(* IEC 61131-3 sources: JingjiangArm/moonboxpro_arm_8.4/Application/Application/任务列表/ExtTask/动作处理/工艺辅助/冷风, 2 files *)

(* ---- KS_ReCfgCoolBlowerIO.st ---- *)
(*@CES
Name=KS_ReCfgCoolBlowerIO
Type=FunctionBlock
TypeGuid=6f9dac99-8de1-4efc-8465-68ac443b7d08
Guid=0f7b114d-d936-480a-be34-fd41a916f68a
HasDeclaration=True
HasImplementation=True
*)
{DECLARATION}
FUNCTION KS_ReCfgCoolBlowerIO : bool
VAR_INPUT
	i_xInput				: BOOL;(*输入重新分配*)
	i_xOutput				: BOOL;(*输出重新分配*)
	i_xCoolBlowerFlag		: BOOL;(*全体冷风启动标志*)
	i_iGrpAxisNum_Pu		:INT ;
	i_aiGrpAxisList			: ARRAY [1..MAX_UNIT_NUM] OF INT;(*系的轴列表*)
	i_paxAxisStartEn		: POINTER TO ARRAY [1..MAX_UNIT_NUM] OF BOOL;(*轴启动使能|有效后按钮开关才能起作用*)
	i_paxStartKnob			: POINTER TO ARRAY [1..MAX_UNIT_NUM] OF BOOL;(*全体启动,每个轴旋钮输入*)
	i_paxStartOrStopBtn		: POINTER TO ARRAY [1..MAX_UNIT_NUM] OF BOOL;(*单轴的启动停止按钮*)
	i_paxNeedStop			: POINTER TO ARRAY [1..MAX_UNIT_NUM] OF BOOL;(*单轴需要停止标志*)
	i_paxAxisStarted		: POINTER TO ARRAY [1..MAX_UNIT_NUM] OF BOOL;(*单个轴的启动输出标志|实际处于启动状态，																		可以根据i_paxNeedStop这个变量控制实际输出*)
	i_axCoolBlower			:ARRAY [1..MAX_UNIT_NUM] OF BOOL;
	i_axCoolBlower_Button			:ARRAY [1..MAX_UNIT_NUM] OF BOOL;
	i_paxLamp_CoolBlower			:POINTER TO ARRAY [1..MAX_UNIT_NUM] OF BOOL;
	i_paxRel_CoolBlower			:POINTER TO ARRAY [1..MAX_UNIT_NUM] OF BOOL;
	i_paxLamp_AllCoolBlower		:POINTER TO ARRAY [1..MAX_UNIT_NUM] OF BOOL;
	i_pxLamp_AllCoolBlower		: POINTER TO BOOL;

END_VAR
VAR_OUTPUT

END_VAR
VAR
	iUnitId: INT;
	iN: INT;
END_VAR

{IMPLEMENTATION}
IF i_paxAxisStartEn<>0 AND
	i_paxStartKnob<>0 AND
	i_paxNeedStop<>0 AND
 	i_paxStartOrStopBtn<>0 AND
	i_paxAxisStarted<>0  THEN
	IF i_xInput THEN
		FOR iN:=1 TO MAX_UNIT_NUM  BY 1 DO
			i_paxStartKnob^[iN]:=FALSE;
			i_paxStartOrStopBtn^[iN]:=FALSE;
			i_paxNeedStop^[iN]:=FALSE;
			i_paxAxisStartEn^[iN]:=FALSE;
		END_FOR

		FOR iN:=1 TO i_iGrpAxisNum_Pu  BY 1 DO
			iUnitId:=i_aiGrpAxisList[iN];
			IF iUnitId>0 AND iUnitId<= MAX_UNIT_NUM THEN
			i_paxStartKnob^[iUnitId]:=i_axCoolBlower[iUnitId];
			i_paxStartOrStopBtn^[iUnitId]:=i_axCoolBlower_Button[iUnitId];
			i_paxNeedStop^[iUnitId]:=FALSE;
			i_paxAxisStartEn^[iUnitId]:=TRUE; (*2024.3.14.165139*)
			END_IF
		END_FOR
	ELSIF i_xOutput THEN
		FOR iN:=1 TO i_iGrpAxisNum_Pu  BY 1 DO
			(*输出到牵引，*)

				iUnitId:=i_aiGrpAxisList[iN];
				IF iUnitId>0 AND iUnitId <= MAX_UNIT_NUM THEN(*输出循环到收牵，这样热风输出灯就可以配到收牵上了|2020.1.9.094955*)
					i_paxLamp_CoolBlower^[iUnitId]:=i_paxAxisStarted^[iUnitId];
					i_paxRel_CoolBlower^[iUnitId]:=i_paxAxisStarted^[iUnitId];
					i_paxLamp_AllCoolBlower^[iUnitId]:=i_xCoolBlowerFlag;
				END_IF

		END_FOR

	END_IF
END_IF

(* ---- KS_FB_GrpCoolBlowerCtrl.st ---- *)
(*@CES
Name=KS_FB_GrpCoolBlowerCtrl
Type=FunctionBlock
TypeGuid=6f9dac99-8de1-4efc-8465-68ac443b7d08
Guid=1cc9b71b-01ee-4c63-826f-1c195b3708a6
HasDeclaration=True
HasImplementation=True
*)
{DECLARATION}
FUNCTION_BLOCK KS_FB_GrpCoolBlowerCtrl
(*2020.10.14.090348重新处理*)
VAR_INPUT
	i_xEn: BOOL;
	i_iGrpId : INT;
	i_iAxisId_If: INT;
	i_iAxisId_Of: INT;
	i_iGrpAxisNum_Pu: INT; (*色组轴数*)
	i_aiGrpAxisList: ARRAY [1..MAX_UNIT_NUM] OF INT; (*系的轴列表*)
	i_pstStEvtReq:POINTER TO StEvtReq;
	i_xCoolBlowerByKnob:BOOL;(*单轴启动根据旋钮开关标志|用于全体开关控制启动的逻辑|无则不输入*)
	i_xStopCoolBlowerWhenEstop:BOOL;(*急停停止热风标志|有效了和急停关联，无效则不影响*)
	i_iCycleTime_Plc:INT;(*2024.01.22.142933+*)
	i_PastStIOMap_Axis_Extra_FE:  POINTER TO ARRAY [1..MAX_UNIT_NUM] OF StIOMap_Axis_Extra_FE  ;

	i_pastStIOMap_Main_FE	: POINTER TO ARRAY [1..4] OF StIOMap_Main_FE;(*轴io数据区域|*)
END_VAR
VAR_OUTPUT
	o_xEno: BOOL;
	o_iErNo: INT;(*0成功\-1参数无效|*)
	o_xCoolBlowerFlag:BOOL;
END_VAR
VAR
	fbKS_FB_CoolBlowerSys: KS_FB_BlowerFunction;
	axAxisStartKnob: ARRAY [1..MAX_UNIT_NUM] OF BOOL;
	axStartOrStopBtn: ARRAY [1..MAX_UNIT_NUM] OF BOOL;
	axNeedStop: ARRAY [1..MAX_UNIT_NUM] OF BOOL;
	axAxisStarted: ARRAY [1..MAX_UNIT_NUM] OF BOOL;
	axAxisStartEn: ARRAY [1..MAX_UNIT_NUM] OF BOOL;
	xCoolBlowerEn: BOOL;
	iStartedSum: INT;(*启动的轴数*)
	xFlag_Estop_In : BOOL;

	axCoolBlower_In			:ARRAY [1..MAX_UNIT_NUM] OF BOOL;
	axCoolBlower_Button_In			:ARRAY [1..MAX_UNIT_NUM] OF BOOL;

	xCoolBlower_In			: BOOL;
	xCoolBlower_Button_In			: BOOL;

	axLamp_CoolBlower_Out			: ARRAY [1..MAX_UNIT_NUM] OF BOOL;
	axRel_CoolBlower_Out			: ARRAY [1..MAX_UNIT_NUM] OF BOOL;
	axLamp_AllCoolBlower_Out	: ARRAY [1..MAX_UNIT_NUM] OF BOOL;
	xLamp_AllCoolBlower_Out	: BOOL;

	pstStIOMap_Axis_Extra_FE:  POINTER TO  StIOMap_Axis_Extra_FE  ;

	iN: INT;
	iUnitId: INT;(*轴号*)
	iGrp: INT;
END_VAR
{IMPLEMENTATION}
Action_Input();

Action_ActCtl() ;

Action_Output();
